(* IEC 61131-3 sources: Test-Git_ESME26/TestProgettoESME_26.fbsproj/TemplateFullProgrammingFramework_Migration.device.xml.v3^/Plc Logic.plclogic.xml.v3^/Application.application.xml.v3^/TemplateFullProgrammingFramework/Examples/ExampleLeafModule, 6 files *)

(* ---- FC_EtDiagExtExampleLeafModuleToString.fn.st ---- *)
FUNCTION FC_EtDiagExtExampleLeafModuleToString : STRING[80]

VAR_INPUT
	i_etDiagExt : ET_DiagExtExampleLeafModule;
END_VAR

VAR_OUTPUT
	q_etDiag	: GD.ET_Diag := GD.ET_Diag.Ok;
	q_etDiagExt	: ET_DiagExtExampleLeafModule := ET_DiagExtExampleLeafModule.Ok;
END_VAR

VAR
END_VAR

CASE i_etDiagExt OF
	ET_DiagExtExampleLeafModule.Ok:										FC_EtDiagExtExampleLeafModuleToString := 'Ok';
	ET_DiagExtExampleLeafModule.Disabled:								FC_EtDiagExtExampleLeafModuleToString := 'Disabled';
	ET_DiagExtExampleLeafModule.Initializing:							FC_EtDiagExtExampleLeafModuleToString := 'Initializing';
	ET_DiagExtExampleLeafModule.NoOp:									FC_EtDiagExtExampleLeafModuleToString := 'NoOp';
	ET_DiagExtExampleLeafModule.HomingWaitForStart:						FC_EtDiagExtExampleLeafModuleToString := 'HomingWaitForStart';
	ET_DiagExtExampleLeafModule.HomingExecuting:						FC_EtDiagExtExampleLeafModuleToString := 'HomingExecuting';
	ET_DiagExtExampleLeafModule.HomingDone:								FC_EtDiagExtExampleLeafModuleToString := 'HomingDone';
	ET_DiagExtExampleLeafModule.AutoWaitForStart:						FC_EtDiagExtExampleLeafModuleToString := 'AutoWaitForStart';
	ET_DiagExtExampleLeafModule.AutoRunning:							FC_EtDiagExtExampleLeafModuleToString := 'AutoRunning';
	ET_DiagExtExampleLeafModule.Working:								FC_EtDiagExtExampleLeafModuleToString := 'Working';

	ET_DiagExtExampleLeafModule.UnknownDiagExtExampleLeafModule:		FC_EtDiagExtExampleLeafModuleToString := 'UnknownDiagExtExampleLeafModule';
	ET_DiagExtExampleLeafModule.SubModuleAddInterfacesInvalidPointer:	FC_EtDiagExtExampleLeafModuleToString := 'SubModuleAddInterfacesInvalidPointer';
	ET_DiagExtExampleLeafModule.SubModuleConstantRange:					FC_EtDiagExtExampleLeafModuleToString := 'SubModuleConstantRange';
	ET_DiagExtExampleLeafModule.MissingExtInit:							FC_EtDiagExtExampleLeafModuleToString := 'MissingExtInit';
	ET_DiagExtExampleLeafModule.ReactionOffsetRange:					FC_EtDiagExtExampleLeafModuleToString := 'ReactionOffsetRange';
	ET_DiagExtExampleLeafModule.DriveInvalid:							FC_EtDiagExtExampleLeafModuleToString := 'DriveInvalid';

	ET_DiagExtExampleLeafModule.CmdUnknown:								FC_EtDiagExtExampleLeafModuleToString := 'CmdUnknown';
	ET_DiagExtExampleLeafModule.CmdImpossibleOverwrite:					FC_EtDiagExtExampleLeafModuleToString := 'CmdImpossibleOverwrite';
	ET_DiagExtExampleLeafModule.CmdImpossibleState:						FC_EtDiagExtExampleLeafModuleToString := 'CmdImpossibleState';
	ET_DiagExtExampleLeafModule.CmdImpossibleReaction:					FC_EtDiagExtExampleLeafModuleToString := 'CmdImpossibleReaction';

	ET_DiagExtExampleLeafModule.AsyncStop:								FC_EtDiagExtExampleLeafModuleToString := 'AsyncStop';
	ET_DiagExtExampleLeafModule.SyncStopEL:								FC_EtDiagExtExampleLeafModuleToString := 'SyncStopEL';
	ET_DiagExtExampleLeafModule.SyncStopEH:								FC_EtDiagExtExampleLeafModuleToString := 'SyncStopEH';
	ET_DiagExtExampleLeafModule.StopEndOfCycle:							FC_EtDiagExtExampleLeafModuleToString := 'StopEndOfCycle';

	ET_DiagExtExampleLeafModule.DriveFatalException:					FC_EtDiagExtExampleLeafModuleToString := 'DriveFatalException';
	ET_DiagExtExampleLeafModule.DriveException:							FC_EtDiagExtExampleLeafModuleToString := 'DriveException';
	ET_DiagExtExampleLeafModule.DriveWarning:							FC_EtDiagExtExampleLeafModuleToString := 'DriveWarning';

	ET_DiagExtExampleLeafModule.UnknownState:							FC_EtDiagExtExampleLeafModuleToString := 'UnknownState';
	ET_DiagExtExampleLeafModule.UnknownCmd:								FC_EtDiagExtExampleLeafModuleToString := 'UnknownCmd';
	ET_DiagExtExampleLeafModule.RandomException:						FC_EtDiagExtExampleLeafModuleToString := 'RandomException';

	ET_DiagExtExampleLeafModule.CurrentStandardItfInvalidPointer:		FC_EtDiagExtExampleLeafModuleToString := 'CurrentStandardItfInvalidPointer';
	ET_DiagExtExampleLeafModule.CurrentAddItfInvalidPointer:			FC_EtDiagExtExampleLeafModuleToString := 'CurrentAddItfInvalidPointer';

	ET_DiagExtExampleLeafModule.ParentInvalid:							FC_EtDiagExtExampleLeafModuleToString := 'ParentInvalid';
	ET_DiagExtExampleLeafModule.ParentNotRegistered:					FC_EtDiagExtExampleLeafModuleToString := 'ParentNotRegistered';
	ET_DiagExtExampleLeafModule.MaxNumberOfLoggerPointsExeeded:			FC_EtDiagExtExampleLeafModuleToString := 'MaxNumberOfLoggerPointsExeeded';
	ET_DiagExtExampleLeafModule.UnexpectedDiagExt:						FC_EtDiagExtExampleLeafModuleToString := 'UnexpectedDiagExt';

	ELSE
		FC_EtDiagExtExampleLeafModuleToString := Standard.CONCAT('Unkown ET_DiagExtExampleLeafModule ', UDINT_TO_STRING(i_etDiagExt));

		q_etDiag	:= GD.ET_Diag.InputParameterInvalid;
		q_etDiagExt	:= ET_DiagExtExampleLeafModule.UnknownDiagExtExampleLeafModule;
END_CASE

(* ---- FC_EtExampleLeafModuleCmdToString.fn.st ---- *)
FUNCTION FC_EtExampleLeafModuleCmdToString : STRING[15]
VAR_INPUT
	i_diCmd		: DINT;
END_VAR
VAR_OUTPUT
	q_etDiag	: GD.ET_Diag := GD.ET_Diag.Ok;
	q_etDiagExt	: ET_DiagExtExampleLeafModule := ET_DiagExtExampleLeafModule.Ok;
END_VAR

CASE i_diCMD OF
	ET_ExampleLeafModuleCmd.Homing:
		FC_EtExampleLeafModuleCmdToString := 'Homing';
	ET_ExampleLeafModuleCmd.Auto:
		FC_EtExampleLeafModuleCmdToString := 'Auto';
	ET_ExampleLeafModuleCmd.Stop:
		FC_EtExampleLeafModuleCmdToString := 'Stop';
	ET_ExampleLeafModuleCmd.Start:
		FC_EtExampleLeafModuleCmdToString := 'Start';
	ET_ExampleLeafModuleCmd.Hold:
		FC_EtExampleLeafModuleCmdToString := 'Hold';
	ELSE
		FC_EtExampleLeafModuleCmdToString := CONCAT('Unkown Cmd ', DINT_TO_STRING(i_diCMD));

		q_etDiag := GD.ET_Diag.InputParameterInvalid;
		q_etDiagExt := ET_DiagExtExampleLeafModule.UnknownCmd;
END_CASE

(* ---- FC_EtExampleLeafModuleStateToString.fn.st ---- *)
FUNCTION FC_EtExampleLeafModuleStateToString : STRING[25]
VAR_INPUT
	i_etState	: ET_ExampleLeafModuleState;
END_VAR
VAR_OUTPUT
	q_etDiag	: GD.ET_Diag := GD.ET_Diag.Ok;
	q_etDiagExt	: ET_DiagExtExampleLeafModule := ET_DiagExtExampleLeafModule.Ok;
END_VAR

CASE i_etState OF
	ET_ExampleLeafModuleState.Disabled:
		FC_EtExampleLeafModuleStateToString := 'Disabled';
	ET_ExampleLeafModuleState.Initializing:
		FC_EtExampleLeafModuleStateToString := 'Initializing';
	ET_ExampleLeafModuleState.NoOp:
		FC_EtExampleLeafModuleStateToString := 'NoOp';
	ET_ExampleLeafModuleState.HomingWaitForStart:
		FC_EtExampleLeafModuleStateToString := 'HomingWaitForStart';
	ET_ExampleLeafModuleState.HomingExecuting:
		FC_EtExampleLeafModuleStateToString := 'HomingExecuting';
	ET_ExampleLeafModuleState.HomingDone:
		FC_EtExampleLeafModuleStateToString := 'HomingDone';
	ET_ExampleLeafModuleState.AutoWaitForStart:
		FC_EtExampleLeafModuleStateToString := 'AutoWaitForStart';
	ET_ExampleLeafModuleState.AutoRunning:
		FC_EtExampleLeafModuleStateToString := 'AutoRunning';
	ELSE
		FC_EtExampleLeafModuleStateToString := CONCAT('Unkown State ', UDINT_TO_STRING(i_etState));

		q_etDiag := GD.ET_Diag.InputParameterInvalid;
		q_etDiagExt := ET_DiagExtExampleLeafModule.UnknownState;
END_CASE

(* ---- FC_UpdateExampleLeafModuleAddInterfaceStruct.fn.st ---- *)
FUNCTION FC_UpdateExampleLeafModuleAddInterfaceStruct : BOOL

VAR_INPUT
	i_pdwSubModuleAddInterfaces		: POINTER TO TPL.TYPE_ADDRESS; // change from DWORD to ADDRESS;
	i_udiSubModuleConstant			: UDINT;
END_VAR

VAR_OUTPUT
	q_etDiag						: GD.ET_Diag := GD.ET_Diag.Ok;
	q_etDiagExt						: ET_DiagExtExampleLeafModule := ET_DiagExtExampleLeafModule.Ok;
	q_sMsg							: STRING[80] := '';
END_VAR

VAR_IN_OUT
	iq_stExampleLeafModuleInterface	: ST_ExampleLeafModuleInterface;
END_VAR

VAR
	pdwArrayPos						: POINTER TO TPL.TYPE_ADDRESS; // change from DWORD to ADDRESS;
END_VAR

IF i_pdwSubModuleAddInterfaces = 0 THEN
	q_etDiag	:= GD.ET_Diag.InputParameterInvalid;
	q_etDiagExt	:= ET_DiagExtExampleLeafModule.SubModuleAddInterfacesInvalidPointer;
	q_sMsg		:= '';
ELSIF i_udiSubModuleConstant < 1 THEN
	q_etDiag	:= GD.ET_Diag.InputParameterInvalid;
	q_etDiagExt := ET_DiagExtExampleLeafModule.SubModuleConstantRange;
	q_sMsg		:= '1 <= i_udiSubModuleConstant';
ELSE
	pdwArrayPos := i_pdwSubModuleAddInterfaces + UDINT_TO_DWORD((i_udiSubModuleConstant-1) * SIZEOF(pdwArrayPos^));
	pdwArrayPos^ := ADR(iq_stExampleLeafModuleInterface);
END_IF

(* ---- FB_ExampleLeafModuleController.fb.st ---- *)
FUNCTION_BLOCK FB_ExampleLeafModuleController

VAR_INPUT
	i_xEnable				: BOOL;
END_VAR

VAR_IN_OUT
	iq_stStandardModuleItf	: TPL.ST_StandardModuleInterface;
	iq_stStandardMotionItf	: TPL.ST_StandardMotionInterface;
	iq_stExceptionList		: TPL.ST_ExceptionList;
	iq_stLogDataList		: TPL.ST_LogDataList;
END_VAR

VAR_OUTPUT
	q_xActive				: BOOL;
	q_xReady				: BOOL;
	q_etDiag				: GD.ET_Diag := GD.ET_Diag.Ok;
	q_etDiagExt				: ET_DiagExtExampleLeafModule := ET_DiagExtExampleLeafModule.Disabled;
	q_sMsg					: STRING[80] := '';
END_VAR

VAR
	xEnableFlag				: BOOL;
	udiTmp					: UDINT;
END_VAR

IF i_xEnable AND NOT xEnableFlag THEN
	xEnableFlag	:= TRUE;

	q_xActive	:= TRUE;

	q_etDiag	:= GD.ET_Diag.Ok;
	q_etDiagExt := ET_DiagExtExampleLeafModule.Initializing;
	q_sMsg		:= '';

	IF ((iq_stStandardModuleItf.iq_stExt.udiNumberOfSubModules <> 0) AND
	   ((iq_stStandardModuleItf.iq_stExt.pdwSubModulesAddItf = 0) OR (iq_stStandardModuleItf.iq_stExt.dwSubModulesItf = 0))) THEN

		q_etDiag	:= GD.ET_Diag.ExecutionAborted;
		q_etDiagExt	:= ET_DiagExtExampleLeafModule.MissingExtInit;
		q_sMsg		:= 'Missing call of FC_UpdateExampleLeafModuleAddInterfaceStruct';

		RETURN;
	END_IF

	udiTmp := ET_ExceptionSource.ExampleLeafModule;

	q_xReady := TPL.FC_CheckSubModuleList(	i_dwModuleType		:= UDINT_TO_DWORD(ET_ModuleType.ExampleLeafModule),
											i_udiModuleId		:= iq_stStandardModuleItf.i_udiModuleId,
											i_sModuleName		:= iq_stStandardModuleItf.i_sModuleName,
											i_etSource			:= udiTmp (* Hack around compiler restrictions *),
											iq_stExt			:= iq_stStandardModuleItf.iq_stExt,
											iq_stExceptionList	:= iq_stExceptionList,
											iq_stLogDataList	:= iq_stLogDataList);

	IF NOT q_xReady THEN
		xEnableFlag := FALSE;
	END_IF

ELSIF NOT i_xEnable AND xEnableFlag THEN
	xEnableFlag	:= FALSE;

	(* No actions required, this simple module does not support jogging or any other things the XXXModuleController would have to handle *)
	q_xReady 	:= FALSE;
	q_xActive	:= FALSE;

	q_etDiag	:= GD.ET_Diag.Ok;
	q_etDiagExt	:= ET_DiagExtExampleLeafModule.Disabled;
	q_sMsg		:= '';
END_IF

IF q_xActive AND q_xReady THEN
	(* No actions required, this simple module does not support jogging or any other things the XXXModuleController would have to handle *)
	q_etDiag	:= GD.ET_Diag.Ok;
	q_etDiagExt := ET_DiagExtExampleLeafModule.Working;
	q_sMsg		:= '';
END_IF

(* ---- FB_ExampleLeafModuleVisController.fb.st ---- *)
FUNCTION_BLOCK FB_ExampleLeafModuleVisController

VAR_INPUT
	i_xEnable								: BOOL;
	i_pstMachineStandardItf					: POINTER TO TPL.ST_StandardModuleInterface;
	i_pstCurrentStandardItf					: POINTER TO TPL.ST_StandardModuleInterface;
	i_dwCurrentAddItf						: TPL.TYPE_ADDRESS; // change DWORD to ADDRESS
	i_xUpdateData							: BOOL; (* Signals the selection of another module *)
	i_udiCurrentJogTarget					: UDINT;
END_VAR

VAR_IN_OUT
	iq_stExceptionList				: TPL.ST_ExceptionList;
	iq_stLogDataList	   			: TPL.ST_LogDataList;
END_VAR

VAR_OUTPUT
	q_xActive								: BOOL;
	q_xReady								: BOOL;
	q_etDiag								: GD.ET_Diag := GD.ET_Diag.Ok;
	q_etDiagExt								: ET_DiagExtExampleLeafModule := ET_DiagExtExampleLeafModule.Disabled;
	q_sMsg									: STRING[80] := '';
	q_udiSetAsCurrentModule					: UDINT; (* A moduleID, if <> 0, it is set as the current module *)
	q_udiSetAsJogTarget						: UDINT;
END_VAR

VAR
	xCurrentIsOfMyType						: BOOL;
	pstCurrentExampleLeafModuleInterface	: POINTER TO ST_ExampleLeafModuleInterface;
	stCurrentExampleLeafModuleInterface		: ST_ExampleLeafModuleInterface;
	iPaneSelect								: INT := 1; (* Variable for selecting the active pane *)

	(* Variables to detect user changes in the vis *)
	xInitUserInputs							: BOOL;

	(* list of all example leaf modules in the machine *)
	audiExampleLeafModuleId					: ARRAY[1..c_udiMaxExampleLeafModules] OF UDINT; (* if <> 0, module exists *)
	asExampleLeafModuleName					: ARRAY[1..c_udiMaxExampleLeafModules] OF STRING[80]; (* if <> 0, module exists *)
	udiCountExampleLeafModules				: UDINT;
	udiSetAsCurrentModule					: UDINT;

	(* temporary variable, not to be used after init *)
	apExampleLeafModuleInterface			: ARRAY[1..c_udiMaxExampleLeafModules] OF POINTER TO TPL.ST_StandardModuleInterface;
	udiTmp									: UDINT;
	xEnableFlag								: BOOL;

	(* Variables to detect user changes in the vis *)
	lrPosMax								: LREAL;
END_VAR

VAR CONSTANT
	c_udiMaxExampleLeafModules : UDINT := 10;
END_VAR

q_udiSetAsCurrentModule 	:= 0;
q_udiSetAsJogTarget			:= 0;

(*********************************************************************)

IF i_xEnable AND NOT xEnableFlag THEN
	xEnableFlag := TRUE;

	q_xActive	:= TRUE;

	q_etDiag	:= GD.ET_Diag.Ok;
	q_etDiagExt := ET_DiagExtExampleLeafModule.Initializing;
	q_sMsg		:= '';

	udiCountExampleLeafModules := TPL.FC_GetAllModulesOfType(	i_pstMachineStandardItf	:= i_pstMachineStandardItf,
																i_dwWantedType			:= ET_ModuleType.ExampleLeafModule,
																i_pdwResultSet			:= ADR(apExampleLeafModuleInterface),
																i_udiResultSetSize		:= c_udiMaxExampleLeafModules);
	FOR udiTmp := 1 TO udiCountExampleLeafModules DO
		(* module version check *)
		IF(apExampleLeafModuleInterface[udiTmp]^.q_udiModuleVersion = 1) THEN
			audiExampleLeafModuleId[udiTmp] := apExampleLeafModuleInterface[udiTmp]^.i_udiModuleId;
			asExampleLeafModuleName[udiTmp] := apExampleLeafModuleInterface[udiTmp]^.i_sModuleName;
		END_IF
	END_FOR

	q_xReady	:= TRUE;

	q_etDiag	:= GD.ET_Diag.Ok;
	q_etDiagExt	:= ET_DiagExtExampleLeafModule.Working;
	q_sMsg		:= '';

ELSIF NOT i_xEnable AND xEnableFlag THEN
	xEnableFlag := FALSE;

	q_xActive				:= FALSE;
	q_xReady				:= FALSE;
	q_etDiag				:= GD.ET_Diag.Ok;
	q_etDiagExt				:= ET_DiagExtExampleLeafModule.Disabled;
	q_sMsg					:= '';
	q_udiSetAsCurrentModule	:= 0;
	q_udiSetAsJogTarget		:= 0;
END_IF

IF i_xEnable THEN
	q_udiSetAsCurrentModule := udiSetAsCurrentModule;
	udiSetAsCurrentModule := 0;
END_IF

(*********************************************************************)

IF i_xEnable THEN
	IF i_pstCurrentStandardItf = 0 THEN
		q_xReady := FALSE;
		q_etDiag := GD.ET_Diag.InputParameterInvalid;
		q_etDiagExt := ET_DiagExtExampleLeafModule.CurrentStandardItfInvalidPointer;
		q_sMsg := '';
	ELSIF i_dwCurrentAddItf = 0 THEN
		q_xReady := FALSE;
		q_etDiag := GD.ET_Diag.InputParameterInvalid;
		q_etDiagExt := ET_DiagExtExampleLeafModule.CurrentAddItfInvalidPointer;
		q_sMsg := '';
	ELSE
		q_xReady	:= TRUE;

		q_etDiag	:= GD.ET_Diag.Ok;
		q_etDiagExt	:= ET_DiagExtExampleLeafModule.Working;
		q_sMsg		:= '';

		IF (i_pstCurrentStandardItf^.q_dwModuleType = UDINT_TO_DWORD(ET_ModuleType.ExampleLeafModule)) THEN
			(* Module version check *)
			IF(i_pstCurrentStandardItf^.q_udiModuleVersion = 1) THEN
				pstCurrentExampleLeafModuleInterface := i_dwCurrentAddItf;
				xCurrentIsOfMyType := TRUE;
			END_IF
		ELSE
			pstCurrentExampleLeafModuleInterface := 0;
			xCurrentIsOfMyType := FALSE;
		END_IF

		IF(xCurrentIsOfMyType) THEN
			(* Execute changes requested by user first *)
			IF(NOT xInitUserInputs) THEN
				xInitUserInputs := TRUE;
				(* Ignore values of variables now *)
			ELSE
				(* Detect user changes *)
				IF stCurrentExampleLeafModuleInterface.i_lrPosMax <> lrPosMax THEN
					pstCurrentExampleLeafModuleInterface^.i_lrPosMax := stCurrentExampleLeafModuleInterface.i_lrPosMax;
				END_IF

				(* ... *)
			END_IF
			stCurrentExampleLeafModuleInterface := pstCurrentExampleLeafModuleInterface^;

		ELSE
			;
			(* Reset other flags *)
		END_IF
	END_IF
ELSE
	xCurrentIsOfMyType := FALSE;
END_IF
